ADAPTER AEquipment (* An adapter: one connection from a skill's run (the plug) to its equipment's port (EP_, the socket) that carries a command out and the word that it was played back. Technical: What a skill's run (SKILL_Run, the plug) sends its equipment's port (EP_, the socket): SEND a command; PLAYED comes back when all its phases are out *)
  (* Standard: 61499-2 *)
  (* Version 0.1, 2026-09-28, Project contributors, AAU Smart Production Lab *)
  PACKAGE modlib;
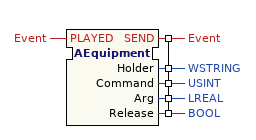
  EVENT_INPUT
    PLAYED; (* All phases of the command were sent *)
  END_EVENT
  EVENT_OUTPUT
    SEND WITH Holder, Command, Arg, Release; (* Send a command to the equipment: its output values, phase by phase *)
  END_EVENT
  VAR_OUTPUT
    Holder : WSTRING; (* Who sends the command *)
    Command : USINT; (* The command's code *)
    Arg : LREAL; (* The command's argument (e.g. a position) *)
    Release : BOOL; (* Give up the equipment after the command *)
  END_VAR
END_ADAPTER
